(* IEC 61131-3 sources: nautilus/website/lessons/b4-counter/start, 1 file *)

(* ---- program.st ---- *)
PROGRAM Counter
VAR
    parcels : CTU;   (* counts, and says when it has reached its preset *)
END_VAR

(* TODO 1: count a parcel each time the eye goes from clear to blocked;
   Reset sets the count back to 0; the preset is 5. *)

(* TODO 2: Count shows the count, and Full is TRUE once 5 have been counted. *)

END_PROGRAM
